Yaskawa INFORM job: SUBPROG.JBI

/JOB
//NAME SUBPROG
//POS
///NPOS 1,0,1,0,0,0
///TOOL 9
///POSTYPE PULSE
///PULSE
C00000=0,0,0
EC00000=0
//INST
<volatile>
///COMM Generated using RoboDK
///ATTR SC,RW
///GROUP1 RB1
NOP
MOVJ C00000 VJ=50.00  +MOVJ EC00000 VJ=100.00
END
